FUNCTION_BLOCK TUNING_TRIGGER (* Select normal control or periodic model tuning; zero interval selects one update *)
  (* Standard: 61499-2 *)
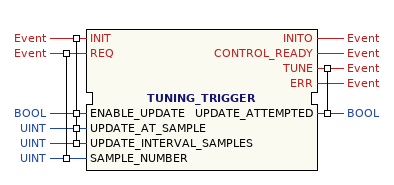
  EVENT_INPUT
    INIT WITH ENABLE_UPDATE, UPDATE_AT_SAMPLE, UPDATE_INTERVAL_SAMPLES;
    REQ WITH SAMPLE_NUMBER;
  END_EVENT
  EVENT_OUTPUT
    INITO;
    CONTROL_READY;
    TUNE WITH UPDATE_ATTEMPTED;
    ERR;
  END_EVENT
  VAR_INPUT
    ENABLE_UPDATE : BOOL;
    UPDATE_AT_SAMPLE : UINT;
    UPDATE_INTERVAL_SAMPLES : UINT;
    SAMPLE_NUMBER : UINT;
  END_VAR
  VAR_OUTPUT
    UPDATE_ATTEMPTED : BOOL;
  END_VAR
  VAR
    ENABLED : BOOL;
    TARGET_SAMPLE : UINT;
    INTERVAL_SAMPLES : UINT;
    LAST_UPDATE_SAMPLE : UINT;
    DUE : BOOL;
    VALID : BOOL;
  END_VAR
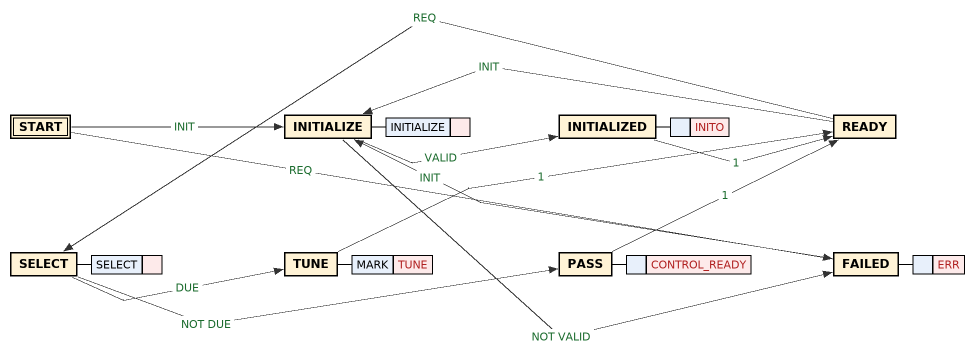
  EC_STATES
    START;
    INITIALIZE : INITIALIZE;
    INITIALIZED : -> INITO;
    READY;
    SELECT : SELECT;
    TUNE : MARK -> TUNE;
    PASS : -> CONTROL_READY;
    FAILED : -> ERR;
  END_STATES
  EC_TRANSITIONS
    START TO INITIALIZE := INIT;
    READY TO INITIALIZE := INIT;
    FAILED TO INITIALIZE := INIT;
    START TO FAILED := REQ;
    INITIALIZE TO INITIALIZED := VALID;
    INITIALIZE TO FAILED := NOT VALID;
    INITIALIZED TO READY := 1;
    READY TO SELECT := REQ;
    SELECT TO TUNE := DUE;
    SELECT TO PASS := NOT DUE;
    TUNE TO READY := 1;
    PASS TO READY := 1;
  END_TRANSITIONS
  ALGORITHM INITIALIZE IN ST:
ENABLED := ENABLE_UPDATE;
TARGET_SAMPLE := UPDATE_AT_SAMPLE;
INTERVAL_SAMPLES := UPDATE_INTERVAL_SAMPLES;
LAST_UPDATE_SAMPLE := 0;
UPDATE_ATTEMPTED := FALSE;
VALID := (NOT ENABLED) OR (TARGET_SAMPLE > 0);
  END_ALGORITHM
  ALGORITHM SELECT IN ST:
DUE := ENABLED AND (NOT UPDATE_ATTEMPTED) AND (SAMPLE_NUMBER = TARGET_SAMPLE);
IF ENABLED AND UPDATE_ATTEMPTED AND (INTERVAL_SAMPLES > 0) AND (SAMPLE_NUMBER >= LAST_UPDATE_SAMPLE) THEN
    DUE := (SAMPLE_NUMBER - LAST_UPDATE_SAMPLE) >= INTERVAL_SAMPLES;
END_IF;
  END_ALGORITHM
  ALGORITHM MARK IN ST:
UPDATE_ATTEMPTED := TRUE;
LAST_UPDATE_SAMPLE := SAMPLE_NUMBER;
  END_ALGORITHM
END_FUNCTION_BLOCK
